(* IEC 61131-3 sources: nautilus/devprofile/profiles, 4 files *)

(* ---- abb-drives.st ---- *)
FUNCTION_BLOCK ABB_DRIVES_SIM
(* An ABB drive under the ABB Drives communication profile, as the FENA /
   FMBT-21 manual (3AUA0000093568 Rev E, pp. 91-96) describes it: the
   control word walks the state machine of p. 95, reference 1 (+-20000 =
   +-100 % of the speed scaling) sets the speed through a linear ramp, and
   the status word reports the state. Simplified: one ramp time, no
   supervision limit (ABOVE_LIMIT stays 0), Actual 2 reads 0, and the drive
   is always in remote (REMOTE = 1). *)
VAR_INPUT
  ControlWord : WORD;
  Reference1 : INT;
  Dt : REAL;              (* seconds since the last scan; the plant wires it *)
  Trip : BOOL;            (* hook: the process model trips the drive *)
  RunEnableLost : BOOL;   (* hook: the external Run enable is off *)
  RampS : REAL;           (* hook: seconds from zero to full speed; 0 means 5 *)
  NominalAmps : REAL;     (* hook: motor current at full load; 0 means 10 *)
  Load : REAL;            (* hook: 0..1, the load the process puts on the motor *)
END_VAR
VAR_OUTPUT
  StatusWord : WORD;
  Actual1 : INT;
  Actual2 : INT;
  Current : REAL;
  Running : BOOL;         (* hook: the motor turns *)
  SpeedPct : REAL;        (* hook: speed in % of the speed scaling *)
END_VAR
VAR
  State : INT;            (* 0 SWITCH-ON INHIBITED, 1 NOT READY TO SWITCH ON,
                             2 READY TO SWITCH ON, 3 READY TO OPERATE,
                             4 OPERATION ENABLED, 9 FAULT *)
  Speed : REAL;
  Fault : BOOL;
  PrevReset : BOOL;
  off1 : BOOL; off2 : BOOL; off3 : BOOL; enable : BOOL; remote : BOOL;
  reset : BOOL; rfgOut : BOOL; rfgHold : BOOL; rfgIn : BOOL;
  ramp : REAL; amps : REAL; target : REAL; step : REAL;
END_VAR
off1 := NOT ControlWord.0;
off2 := NOT ControlWord.1;
off3 := NOT ControlWord.2;
enable := ControlWord.3;
rfgOut := ControlWord.4;
rfgHold := ControlWord.5;
rfgIn := ControlWord.6;
reset := ControlWord.7 AND NOT PrevReset;
PrevReset := ControlWord.7;
remote := ControlWord.10;
ramp := RampS;
IF ramp <= 0.0 THEN ramp := 5.0; END_IF;
amps := NominalAmps;
IF amps <= 0.0 THEN amps := 10.0; END_IF;

(* FAULT from any state; RESET (a rising edge of bit 7) clears it once the
   cause is gone, and the drive goes to SWITCH-ON INHIBITED. *)
IF Trip THEN
  Fault := TRUE;
END_IF;
IF Fault AND reset AND NOT Trip THEN
  Fault := FALSE;
  State := 0;
END_IF;

IF Fault THEN
  State := 9;
ELSIF off2 OR off3 THEN
  State := 0;
ELSE
  CASE State OF
    0: IF off1 THEN State := 1; END_IF;
    1: IF off1 AND remote THEN State := 2; END_IF;
    2: IF NOT off1 AND remote THEN State := 3; END_IF;
    3: IF off1 THEN
         State := 2;
       ELSIF enable AND NOT RunEnableLost THEN
         State := 4;
       END_IF;
    4: IF off1 THEN
         State := 2;
       ELSIF NOT enable OR RunEnableLost THEN
         State := 3;
       END_IF;
  END_CASE;
END_IF;

(* The ramp function generator. *)
target := 0.0;
IF State = 4 AND rfgOut AND rfgIn AND remote THEN
  target := INT_TO_REAL(Reference1);
END_IF;
step := 20000.0 * Dt / ramp;
IF Fault OR off2 THEN
  Speed := 0.0;
ELSIF off3 THEN
  step := step * 10.0;
END_IF;
IF State = 4 AND NOT rfgHold THEN
  step := 0.0;
END_IF;
IF Speed < target THEN
  Speed := MIN(Speed + step, target);
ELSIF Speed > target THEN
  Speed := MAX(Speed - step, target);
END_IF;

Running := ABS(Speed) > 1.0;
SpeedPct := Speed / 200.0;
Actual1 := REAL_TO_INT(Speed);
Actual2 := 0;
IF Running THEN
  Current := amps * (0.3 + 0.7 * Load) * ABS(Speed) / 20000.0;
ELSE
  Current := 0.0;
END_IF;

StatusWord := 0;
StatusWord.0 := State >= 2 AND State <= 4;
StatusWord.1 := State >= 3 AND State <= 4;
StatusWord.2 := State = 4;
StatusWord.3 := Fault;
StatusWord.4 := NOT off2;
StatusWord.5 := NOT off3;
StatusWord.6 := State = 0;
StatusWord.8 := State = 4 AND ABS(Speed - target) <= 2000.0;
StatusWord.9 := TRUE;
StatusWord.11 := ControlWord.11;
StatusWord.12 := NOT RunEnableLost;
END_FUNCTION_BLOCK

(* ---- asi-275m.st ---- *)
FUNCTION_BLOCK ASI_275M_SIM
(* A 16-in/16-out relay board: the controller writes one word of relay
   outputs and reads one word of inputs, point n on bit n-1. The relays and
   inputs are hooks for the process model. *)
VAR_INPUT
  Outputs : WORD;
  Input1 : BOOL; Input2 : BOOL; Input3 : BOOL; Input4 : BOOL;
  Input5 : BOOL; Input6 : BOOL; Input7 : BOOL; Input8 : BOOL;
  Input9 : BOOL; Input10 : BOOL; Input11 : BOOL; Input12 : BOOL;
  Input13 : BOOL; Input14 : BOOL; Input15 : BOOL; Input16 : BOOL;
END_VAR
VAR_OUTPUT
  Inputs : WORD;
  Relay1 : BOOL; Relay2 : BOOL; Relay3 : BOOL; Relay4 : BOOL;
  Relay5 : BOOL; Relay6 : BOOL; Relay7 : BOOL; Relay8 : BOOL;
  Relay9 : BOOL; Relay10 : BOOL; Relay11 : BOOL; Relay12 : BOOL;
  Relay13 : BOOL; Relay14 : BOOL; Relay15 : BOOL; Relay16 : BOOL;
END_VAR
Relay1 := Outputs.0;   Relay2 := Outputs.1;   Relay3 := Outputs.2;   Relay4 := Outputs.3;
Relay5 := Outputs.4;   Relay6 := Outputs.5;   Relay7 := Outputs.6;   Relay8 := Outputs.7;
Relay9 := Outputs.8;   Relay10 := Outputs.9;  Relay11 := Outputs.10; Relay12 := Outputs.11;
Relay13 := Outputs.12; Relay14 := Outputs.13; Relay15 := Outputs.14; Relay16 := Outputs.15;
Inputs := 0;
Inputs.0 := Input1;   Inputs.1 := Input2;   Inputs.2 := Input3;   Inputs.3 := Input4;
Inputs.4 := Input5;   Inputs.5 := Input6;   Inputs.6 := Input7;   Inputs.7 := Input8;
Inputs.8 := Input9;   Inputs.9 := Input10;  Inputs.10 := Input11; Inputs.11 := Input12;
Inputs.12 := Input13; Inputs.13 := Input14; Inputs.14 := Input15; Inputs.15 := Input16;
END_FUNCTION_BLOCK

(* ---- fdc-mct4.st ---- *)
FUNCTION_BLOCK MCT4_SIM
(* An FDC MCT4's loop 1 (MCT4 4.3 User Manual Rev. G, App. A.1): a PI loop
   driving a burner's firing rate, over a first-order thermal model. Heat
   enters only while the burner manager reports a flame. In manual (Manual
   Override bit 0) the output is what the controller wrote to %Out. *)
VAR_INPUT
  AlarmReset : UINT;
  ManualOverride : WORD;
  SystemEvents : WORD;
  Loop1SP : INT;
  Dt : REAL;
  FlameOn : BOOL;       (* hook: the burner manager has a flame *)
  SensorBreak : BOOL;   (* hook: the loop's thermocouple breaks *)
  Ambient : REAL;       (* hook: temperature with no heat; 0 means 70 *)
  HeatRate : REAL;      (* hook: degrees per second at 100 % with a flame; 0 means 5 *)
  LossRate : REAL;      (* hook: share of (PV - ambient) lost per second; 0 means 0.01 *)
END_VAR
VAR_IN_OUT
  Loop1Out : REAL;      (* %Out: the controller's in manual, the loop's in auto *)
END_VAR
VAR_OUTPUT
  OfflineBusy : UINT;
  LoopErrorStatus : WORD;
  AlarmStatus1 : WORD;
  Loop1PV : INT;
  Loop1Status : WORD;
  Loop1Error : UINT;
  Temperature : REAL;   (* hook: the modelled temperature *)
END_VAR
VAR
  pv : REAL;
  started : BOOL;
  integ : REAL;
  e : REAL;
  amb : REAL;
  heat : REAL;
  loss : REAL;
  manual : BOOL;
END_VAR
amb := Ambient;
IF amb = 0.0 THEN amb := 70.0; END_IF;
heat := HeatRate;
IF heat <= 0.0 THEN heat := 5.0; END_IF;
loss := LossRate;
IF loss <= 0.0 THEN loss := 0.01; END_IF;
IF NOT started THEN
  pv := amb;
  started := TRUE;
END_IF;

manual := ManualOverride.0;
IF manual THEN
  Loop1Out := LIMIT(0.0, Loop1Out, 100.0);
  integ := Loop1Out;   (* bumpless back to auto *)
ELSIF SensorBreak THEN
  Loop1Out := 0.0;     (* no measurement, no heat *)
ELSE
  e := INT_TO_REAL(Loop1SP) - pv;
  integ := LIMIT(0.0, integ + 0.2 * e * Dt, 100.0);
  Loop1Out := LIMIT(0.0, 4.0 * e + integ, 100.0);
END_IF;

IF FlameOn THEN
  pv := pv + heat * Loop1Out / 100.0 * Dt;
END_IF;
pv := pv - loss * (pv - amb) * Dt;

Temperature := pv;
Loop1PV := REAL_TO_INT(pv);
Loop1Error := 0;
IF SensorBreak THEN
  Loop1Error := 39;
END_IF;
LoopErrorStatus := 0;
LoopErrorStatus.0 := SensorBreak;
Loop1Status := 0;
Loop1Status.2 := NOT manual;   (* Static Mode: no automatic program *)
Loop1Status.4 := manual;       (* Manual Mode *)
AlarmStatus1 := 0;
OfflineBusy := 0;
END_FUNCTION_BLOCK

(* ---- ifm-al1590.st ---- *)
FUNCTION HEX4 : STRING
(* A word as the four upper-case hex digits an ifm master's pdin carries. *)
VAR_INPUT
  V : UINT;
END_VAR
VAR
  i : INT;
  d : UINT;
  w : UINT;
END_VAR
HEX4 := '';
w := V;
FOR i := 1 TO 4 DO
  d := w MOD 16;
  w := w / 16;
  CASE d OF
    0: HEX4 := CONCAT('0', HEX4);
    1: HEX4 := CONCAT('1', HEX4);
    2: HEX4 := CONCAT('2', HEX4);
    3: HEX4 := CONCAT('3', HEX4);
    4: HEX4 := CONCAT('4', HEX4);
    5: HEX4 := CONCAT('5', HEX4);
    6: HEX4 := CONCAT('6', HEX4);
    7: HEX4 := CONCAT('7', HEX4);
    8: HEX4 := CONCAT('8', HEX4);
    9: HEX4 := CONCAT('9', HEX4);
    10: HEX4 := CONCAT('A', HEX4);
    11: HEX4 := CONCAT('B', HEX4);
    12: HEX4 := CONCAT('C', HEX4);
    13: HEX4 := CONCAT('D', HEX4);
    14: HEX4 := CONCAT('E', HEX4);
  ELSE
    HEX4 := CONCAT('F', HEX4);
  END_CASE;
END_FOR;
END_FUNCTION

FUNCTION_BLOCK IFM_AL1590_SIM
(* Each port's pdin, as hex text, from a word the process model sets. *)
VAR_INPUT
  Port1_Word : UINT; Port2_Word : UINT; Port3_Word : UINT; Port4_Word : UINT;
  Port5_Word : UINT; Port6_Word : UINT; Port7_Word : UINT; Port8_Word : UINT;
END_VAR
VAR_OUTPUT
  Port1_Pdin : STRING; Port2_Pdin : STRING; Port3_Pdin : STRING; Port4_Pdin : STRING;
  Port5_Pdin : STRING; Port6_Pdin : STRING; Port7_Pdin : STRING; Port8_Pdin : STRING;
END_VAR
Port1_Pdin := HEX4(Port1_Word); Port2_Pdin := HEX4(Port2_Word);
Port3_Pdin := HEX4(Port3_Word); Port4_Pdin := HEX4(Port4_Word);
Port5_Pdin := HEX4(Port5_Word); Port6_Pdin := HEX4(Port6_Word);
Port7_Pdin := HEX4(Port7_Word); Port8_Pdin := HEX4(Port8_Word);
END_FUNCTION_BLOCK
